Yaskawa INFORM job: DEMO_C_PLACE.JBI

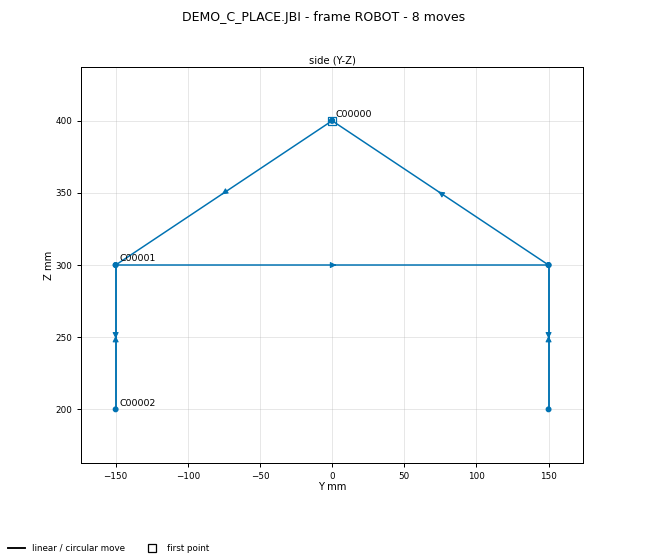
[picture p0: tool path of DEMO_C_PLACE.JBI in frame ROBOT, 8 of 8 moves have a stored position in this frame; points joined in program order, loops and branches not executed]
/JOB
//NAME DEMO_C_PLACE
//POS
///NPOS 8,0,0,0,0,0
///TOOL 0
///POSTYPE ROBOT
///RECTAN
///RCONF 0,0,0,0,0,0,0,0
C00000=400.000,0.000,400.000,180.00,0.00,0.00
C00001=400.000,-150.000,300.000,180.00,0.00,0.00
C00002=400.000,-150.000,200.000,180.00,0.00,0.00
C00003=400.000,-150.000,300.000,180.00,0.00,0.00
C00004=400.000,150.000,300.000,180.00,0.00,0.00
C00005=400.000,150.000,200.000,180.00,0.00,0.00
C00006=400.000,150.000,300.000,180.00,0.00,0.00
C00007=400.000,0.000,400.000,180.00,0.00,0.00
//INST
///DATE 2026/11/02 18:30
///ATTR SC,RW
///GROUP1 RB1
NOP
'SYNTHETIC DEMO JOB - NOT A REAL ROBOT JOB
MOVL C00000 V=200.0
MOVL C00001 V=200.0
MOVL C00002 V=50.0 PL=0
DOUT OT#(1) ON
TIMER T=0.50
MOVL C00003 V=50.0 PL=0
MOVL C00004 V=200.0 PL=0
MOVL C00005 V=50.0 PL=0
TIMER T=3.00
DOUT OT#(1) OFF
TIMER T=0.50
MOVL C00006 V=50.0 PL=0
MOVL C00007 V=200.0
END
